(* Logix 5000 project; controller _1407974_PSG_7315 vendor 1 type 14 code 154 rev 20.11; software revision 20.06 *)
// S/O:1407974
// MODEL: PSG P7315

TASK MainTask (continuous, watchdog 500 ms) : MainProgram

MODULES
   Local : vendor 1 type 14 code 154 (PointIO 0, rev 20.11)
      Delta_V : 1756-ENBT (Ethernet 192.168.1.1, rev 3.1)
      Remote : vendor 1 type 12 code 132 (Ethernet 192.168.1.51, rev 4.10, Output RPI 20 ms)
         RTD_In_Module : vendor 1 type 115 code 125 (ArmorPoint 2, rev 3.4, Input RPI 50 ms)
         DI_1_Module : vendor 1 type 7 code 201 (ArmorPoint 1, rev 3.22, Input RPI 50 ms)
         DO_Module : vendor 1 type 7 code 209 (ArmorPoint 3, rev 3.22, Output RPI 50 ms)
         AO_Module : vendor 1 type 115 code 127 (ArmorPoint 4, rev 3.4, Output RPI 80 ms)
      Local_AI_Slot_2 : 1734-IE2C (PointIO 2, rev 3.1, Input RPI 80 ms)
       : vendor 1 type 115 code 211 (PointIO 3, rev 3.1, Output RPI 80 ms)
      Discrete_IO : Embedded (PointIO 1, rev 20.11, Output RPI 20 ms)
END_MODULES

TYPE Analog_Input :
STRUCT
   Raw : REAL;
   Scaled : REAL;
   Fault : BOOL;
   Under_Range : BOOL;
   Over_Range : BOOL;
   Control_Set_Point : REAL;
   Alarm_Low_Set_Point : REAL;
   Alarm_High_Set_Point : REAL;
   Temp_Set_Point : REAL;
   Tieback : REAL;
   SCP : SCP;
   EU_Low : REAL;
   EU_hi : REAL;
   PID : PID;
   Low_Stpt : REAL;
   Low_Low_Stpt : REAL;
   High_Stpt : REAL;
   High_High_Stpt : REAL;
   Ana_Out : Analog_Output;
END_STRUCT
END_TYPE

TYPE Analog_Output :
STRUCT
   Scaled : REAL;
   Manual : REAL;
   Fault : BOOL;
   Raw : REAL;
   SCP : SCP;
   ManSCP : SCP;
   Set_Point_Entry : OIT_Set_Point_Entry;
END_STRUCT
END_TYPE

TYPE AW :
STRUCT
   Network_Ack : INT[2];
   Network_Ack_ONS : INT[2];
   Network_Ack_Handshake : INT[2];
   Network_Ack_Latch : INT[2];
   Network_Ack_All_Latch : BOOL;
   Remote_Ack_All : INT;
   Network_Alarm_Ack : INT[2];
   OIT_Ack : INT[2];
   Latch_Bit : INT[2];
   Ack : INT[2];
   No_Active_Alarms : BOOL;
   No_Active_Warnings : BOOL;
   Silence : INT[2];
   All_Alarms_Acknowledged : BOOL;
   All_Warnings_Acknowledged : BOOL;
   Alarms_Silenced : BOOL;
   Warnings_Silenced : BOOL;
   OIT_Silence_PB : Push_Button;
   Alarm_Silence_Latch : BOOL;
   Warning_Silence_Latch : BOOL;
END_STRUCT
END_TYPE

TYPE Date_Time :
STRUCT
   Set_Push_Button : BOOL;
   Handshake : BOOL;
END_STRUCT
END_TYPE

TYPE Discrete_Out :
STRUCT
   Activate : BOOL;
   Maint_Latch : Latched_Push_Button;
END_STRUCT
END_TYPE

TYPE OIT_Connections :
STRUCT
   Current_Minute : DINT;
   Update : BOOL;
   Current_Screen : DINT;
   Previous_Minute : DINT;
END_STRUCT
END_TYPE

TYPE OIT_Message :
STRUCT
   Operational_Mode : INT;
   Operational_Step_State : INT;
   Information_Message_Number : INT;
   Feed_Water_Pump_Status : INT;
   Low_Level_Swtitch_Status : INT;
   Hi_Hi_Level_Switch_Status : INT;
   Pure_Steam_Temp_Status : INT;
   Pure_Steam_Conductivity_Status : INT;
   Alarm_Warning_Status : INT;
END_STRUCT
END_TYPE

TYPE OIT_Popup :
STRUCT
   Call : BOOL;
   Called : BOOL;
   Timer : TIMER;
   Close : BOOL;
END_STRUCT
END_TYPE

TYPE OIT_Set_Point_Entry :
STRUCT
   OIT_Enter : Push_Button;
   OIT_Set_Point_Buffer : REAL;
END_STRUCT
END_TYPE

TYPE Push_Button :
STRUCT
   Push_Button : BOOL;
   Indicator : BOOL;
   One_Shot : BOOL;
   Handshake : BOOL;
END_STRUCT
END_TYPE

TYPE Unit_Status :
STRUCT
   ON : BOOL;
   OFF : BOOL;
   READY : BOOL;
   FILLING : BOOL;
   HEATING : BOOL;
   RUNNING : BOOL;
   COOLING : BOOL;
   MAINTENANCE : BOOL;
END_STRUCT
END_TYPE

ADD_ON_INSTRUCTION Latched_Push_Button   (* revision 1.0 *)
VAR_INPUT
   OIT_Momentary_PB : BOOL; {required}
END_VAR
VAR_OUTPUT
   OIT_Status : BOOL; {access Read Only, required}
END_VAR
VAR
   OIT_Toggle_ONS : BOOL;
   OIT_Select_ONS : BOOL;
END_VAR

ROUTINE Logic   (* ladder *)
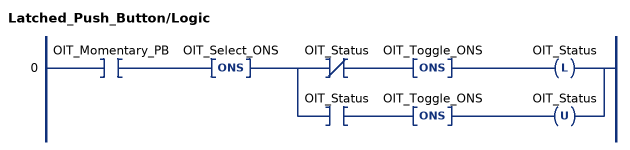
   0: XIC(OIT_Momentary_PB)ONS(OIT_Select_ONS)[XIO(OIT_Status) ONS(OIT_Toggle_ONS) OTL(OIT_Status) ,XIC(OIT_Status) ONS(OIT_Toggle_ONS) OTU(OIT_Status) ];
END_ROUTINE
END_ADD_ON_INSTRUCTION

ADD_ON_INSTRUCTION SCP   (* revision 1.0, vendor Rockwell Automation *)
VAR_INPUT
   Input : REAL; {required}
   InputMin : REAL; {required}
   InputMax : REAL; {required}
   ScaledMin : REAL; {required}
   ScaledMax : REAL; {required}
END_VAR
VAR_OUTPUT
   Output : REAL; {access Read Only, required}
END_VAR
VAR
   Temp4 : REAL;
   Temp3 : REAL;
   Temp2 : REAL;
   Temp1 : REAL;
   Offset : REAL;
   Rate : REAL;
   Out : REAL;
END_VAR

ROUTINE Logic   (* ladder *)
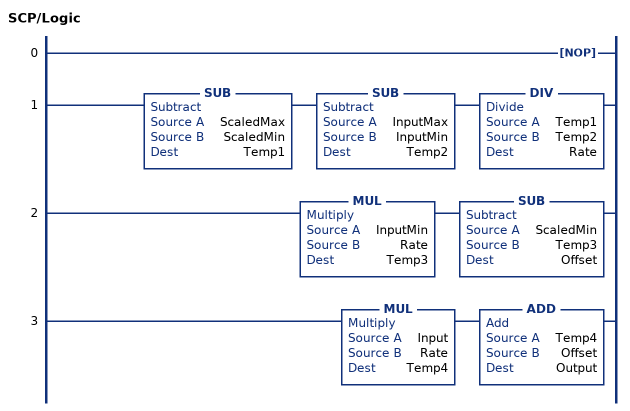
   0: NOP();
   1: SUB(ScaledMax,ScaledMin,Temp1)SUB(InputMax,InputMin,Temp2)DIV(Temp1,Temp2,Rate);
   2: MUL(InputMin,Rate,Temp3)SUB(ScaledMin,Temp3,Offset);
   3: MUL(Input,Rate,Temp4)ADD(Temp4,Offset,Output);
END_ROUTINE
END_ADD_ON_INSTRUCTION

VAR_GLOBAL   (* controller tags *)
   AI_L_2_0_Pure_Steam_Conductivity : Analog_Input := (Raw := 9171.0, Scaled := 0.8994354, Alarm_High_Set_Point := 1.2, SCP.Input := 9171.0, SCP.InputMin := 3277.0, SCP.InputMax := 16383.0, SCP.ScaledMax := 2.0, SCP.Output := 0.8994354);
   AI_L_2_1_FW_Press_Low_Warning : OIT_Set_Point_Entry := (OIT_Set_Point_Buffer := 5.0);
   AI_L_2_1_FW_Pressure : Analog_Input := (Raw := 3321.0, Scaled := 0.5035858, Control_Set_Point := 80.0, Alarm_High_Set_Point := 2.0, Temp_Set_Point := 80.0, SCP.Input := 3321.0, SCP.InputMin := 3277.0, SCP.InputMax := 16383.0, SCP.ScaledMax := 150.0, SCP.Output := 0.5035858, Low_Stpt := 5.0);
   AI_R_2_0_Pure_Steam_Temperature : Analog_Input := (Scaled := 139.6, Control_Set_Point := 140.0, Alarm_Low_Set_Point := 102.0, Alarm_High_Set_Point := 176.0, Temp_Set_Point := 140.0);
   AI_R_2_1_Cond_Pure_Steam_Temperature : Analog_Input := (Scaled := 99.9, Alarm_High_Set_Point := 99.0);
   Alarm_Emergency_Stop : ALIAS FOR Alarms_Warnings.Latch_Bit[0].0;
   Alarm_Emergency_Stop_Ack : ALIAS FOR Alarms_Warnings.Ack[0].0;
   Alarm_Pure_Steam_High_Temp_Timer : TIMER := (PRE := 60000);
   Alarm_Pure_Steam_High_Temperature : ALIAS FOR Alarms_Warnings.Latch_Bit[0].4;
   Alarm_Pure_Steam_High_Temperature_Ack : ALIAS FOR Alarms_Warnings.Ack[0].4;
   Alarm_Pure_Steam_Temp_Error_Timer : TIMER := (PRE := 5000);
   Alarm_Pure_Steam_Temp_Input_Error : ALIAS FOR Alarms_Warnings.Latch_Bit[0].5;
   Alarm_Pure_Steam_Temp_Input_Error_Ack : ALIAS FOR Alarms_Warnings.Ack[0].5;
   Alarm_Rupture_Disk_Failure : ALIAS FOR Alarms_Warnings.Latch_Bit[0].1;
   Alarm_Rupture_Disk_Failure_Timer : TIMER := (PRE := 750);
   Alarm_Rupture_Disk_Faiure_Ack : ALIAS FOR Alarms_Warnings.Ack[0].1;
   Alarm_Separator_High_Level : ALIAS FOR Alarms_Warnings.Latch_Bit[0].2;
   Alarm_Separator_High_Level_Ack : ALIAS FOR Alarms_Warnings.Ack[0].2;
   Alarm_Separator_High_Level_Timer : TIMER := (PRE := 120000);
   Alarm_Separator_Low_Level : ALIAS FOR Alarms_Warnings.Latch_Bit[0].3;
   Alarm_Separator_Low_Level_Ack : ALIAS FOR Alarms_Warnings.Ack[0].3;
   Alarm_Separator_Low_Level_Timer_A : TIMER := (PRE := 600000);
   Alarm_Separator_Low_Level_Timer_B : TIMER := (PRE := 60000);
   Alarms_Warnings : AW := (Network_Ack[1] := 32, Network_Ack_Handshake[0] := 1, Network_Ack_Handshake[1] := 1, Latch_Bit[1] := 2#0000_0000_0000_0001, No_Active_Alarms := 1, All_Alarms_Acknowledged := 1, Alarms_Silenced := 1);
   AO_L_3_0_VFD_SPEED : Analog_Output := (Scaled := 100.0, Manual := 100.0, Raw := 100.0);
   AO_L_3_1_Available : Analog_Output := (SCP.InputMax := 100.0, SCP.ScaledMin := 3277.0, SCP.ScaledMax := 16383.0, SCP.Output := 3277.0, ManSCP.InputMax := 100.0, ManSCP.ScaledMin := 3277.0, ManSCP.ScaledMax := 16383.0, ManSCP.Output := 3277.0);
   AO_L_3_2_Available : Analog_Output := (SCP.InputMax := 100.0, SCP.ScaledMin := 3277.0, SCP.ScaledMax := 16383.0, SCP.Output := 3277.0, ManSCP.InputMax := 100.0, ManSCP.ScaledMin := 3277.0, ManSCP.ScaledMax := 16383.0, ManSCP.Output := 3277.0);
   AO_L_3_3_Available : Analog_Output := (SCP.InputMax := 100.0, SCP.ScaledMin := 3277.0, SCP.ScaledMax := 16383.0, SCP.Output := 3277.0, ManSCP.InputMax := 100.0, ManSCP.ScaledMin := 3277.0, ManSCP.ScaledMax := 16383.0, ManSCP.Output := 3277.0);
   AO_R_4_0_Pure_Steam_Temperature : Analog_Output := (Raw := 54.780636);
   AO_R_4_1_Available : Analog_Output := (SCP.InputMax := 100.0, SCP.ScaledMax := 16383.0, ManSCP.InputMax := 100.0, ManSCP.ScaledMin := 3277.0, ManSCP.ScaledMax := 16383.0, ManSCP.Output := 3277.0);
   Calculated_CV_Max_Value : REAL := 100.0;
   Clean_Steam_Gen_Binary_Data : INT := 8;
   Clean_Steam_Gen_Data : REAL[2] := ([0] := 22.3, [1] := 0.32427895);
   Clean_Steam_Gen_Data3 : INT := 8;
   Cond_Pure_Steam_Conductivity_High : BOOL;
   Cond_Pure_Steam_Hi_Cond_Set_Point_Entry : OIT_Set_Point_Entry := (OIT_Set_Point_Buffer := 1.2);
   Cond_Pure_Steam_Hi_Temp_Set_Point_Entry : OIT_Set_Point_Entry := (OIT_Set_Point_Buffer := 99.0);
   Cond_Pure_Steam_Quality_OK_Latch : BOOL;
   Condensed_Pure_Steam_Warrnings_Disabled : Latched_Push_Button := (OIT_Status := 1);
   Conductivity_Analzyer_Warmup_Delay_Timer : TIMER := (PRE := 600000);
   Cooling_State_Latch_Timer : TIMER := (PRE := 30000, EN := 1, DN := 1);
   Cooling_Status_Debounce_Timer : TIMER := (PRE := 5000);
   DI_L_1_0_Emergency_Stop_Relay : ALIAS FOR DI_Local_1.0;
   DI_L_1_10_Available : ALIAS FOR DI_Local_1.10;
   DI_L_1_11_Available : ALIAS FOR DI_Local_1.11;
   DI_L_1_12_Available : ALIAS FOR DI_Local_1.12;
   DI_L_1_13_Available : ALIAS FOR DI_Local_1.13;
   DI_L_1_14_Feed_Water_Pump_Auto : ALIAS FOR DI_Local_1.14;
   DI_L_1_15_Feed_Water_Pump_Manual : ALIAS FOR DI_Local_1.15;
   DI_L_1_1_Feed_Water_Pump_Aux : ALIAS FOR DI_Local_1.1;
   DI_L_1_2_Pure_Steam_Analyzer_Fault : ALIAS FOR DI_Local_1.2;
   DI_L_1_3_Feed_Water_Analyzer_Fault : ALIAS FOR DI_Local_1.3;
   DI_L_1_4_Available : ALIAS FOR DI_Local_1.4;
   DI_L_1_5_Available : ALIAS FOR DI_Local_1.5;
   DI_L_1_6_Available : ALIAS FOR DI_Local_1.6;
   DI_L_1_7_Available : ALIAS FOR DI_Local_1.7;
   DI_L_1_8_Available : ALIAS FOR DI_Local_1.8;
   DI_L_1_9_Available : ALIAS FOR DI_Local_1.9;
   DI_Local_1 : INT := 7;
   DI_R_1_0_Hi_Hi_Level_LSHH_1950 : ALIAS FOR DI_Remote_1.0;
   DI_R_1_1_Hi_Level_LSH_1950 : ALIAS FOR DI_Remote_1.1;
   DI_R_1_2_Mid_Level_LSM_1950 : ALIAS FOR DI_Remote_1.2;
   DI_R_1_3_Low_Level_LSL_1950 : ALIAS FOR DI_Remote_1.3;
   DI_R_1_4_Air_Low_Pressure_PSL_4030 : ALIAS FOR DI_Remote_1.4;
   DI_R_1_5_Burst_Disk_Sensor_PSH_5820 : ALIAS FOR DI_Remote_1.5;
   DI_R_1_6_Available : ALIAS FOR DI_Remote_1.6;
   DI_R_1_7_Available : ALIAS FOR DI_Remote_1.7;
   DI_Remote_1 : INT := 59;
   DO_L_1_0_Alarm_Relay_Coil : Discrete_Out;
   DO_L_1_0_Alarm_Relay_Out : BOOL;
   DO_L_1_10_Available : Discrete_Out;
   DO_L_1_10_Spare_Out : BOOL;
   DO_L_1_11_Available : Discrete_Out;
   DO_L_1_11_Spare_Out : BOOL;
   DO_L_1_12_Available : Discrete_Out;
   DO_L_1_12_Spare_Out : BOOL;
   DO_L_1_13_Available : Discrete_Out;
   DO_L_1_13_Spare_Out : BOOL;
   DO_L_1_13_VFD_Relay_In : BOOL;
   DO_L_1_14_Feed_Pump_Out : BOOL;
   DO_L_1_14_Feed_Water_Pump_Contactor : Discrete_Out;
   DO_L_1_15_Feed_Pump_Light_Out : BOOL;
   DO_L_1_15_Feed_Water_Pump_On_Light : Discrete_Out;
   DO_L_1_1_Alarm_Horn : Discrete_Out := (Activate := 1);
   DO_L_1_1_Alarm_Horn_Out : BOOL := 1;
   DO_L_1_2_Alarm_Light : Discrete_Out := (Activate := 1);
   DO_L_1_2_Alarm_Light_Out : BOOL := 1;
   DO_L_1_3_Ready_Light : Discrete_Out;
   DO_L_1_3_Ready_Light_Out : BOOL;
   DO_L_1_4_Running_Light : Discrete_Out;
   DO_L_1_4_Running_Light_Out : BOOL;
   DO_L_1_5_Hour_Meter : Discrete_Out;
   DO_L_1_5_Hour_Meter_Out : BOOL;
   DO_L_1_6_Available : Discrete_Out;
   DO_L_1_6_Spare_Out : BOOL;
   DO_L_1_7_Available : Discrete_Out;
   DO_L_1_7_Spare_Out : BOOL;
   DO_L_1_8_Available : Discrete_Out;
   DO_L_1_8_Spare_Out : BOOL;
   DO_L_1_9_Available : Discrete_Out;
   DO_L_1_9_Spare_Out : BOOL;
   DO_Local_1 : INT := 6;
   DO_R_3_0_Pure_Steam_Control_Valve_Out : BOOL;
   DO_R_3_0_Pure_Steam_Temp_Control_YV_4110 : Discrete_Out;
   DO_R_3_1_Pri_Level_Valve_Out : BOOL;
   DO_R_3_1_Primary_Level_Control_YV_4760 : Discrete_Out;
   DO_R_3_2_Sec_Level_Valve_Out : BOOL;
   DO_R_3_2_Secondary_Level_Control_YV_4770 : Discrete_Out;
   DO_R_3_3_Coolant_Shutoff_FCV_3025 : Discrete_Out;
   DO_R_3_3_Coolant_Valve_Out : BOOL;
   DO_R_3_4_Degasser_Vent_Out : BOOL := 1;
   DO_R_3_4_Degasser_Vent_YV_4255 : Discrete_Out := (Activate := 1);
   DO_R_3_5_FDW_TR : Discrete_Out;
   DO_R_3_5_Spare_Out : BOOL;
   DO_R_3_6_Available : Discrete_Out;
   DO_R_3_6_Spare_Out : BOOL;
   DO_R_3_7_Available : Discrete_Out;
   DO_R_3_7_Spare_Out : BOOL;
   DO_Remote_3 : INT := 16;
   F8_0_9 : REAL[10] := ([0] := 139.6, [1] := 0.8994354); {produced, access Read Only}
   F8_50_59 : REAL[10]; {produced}
   Feed_Water_Conductivity_High : BOOL;
   Feed_Water_Pressure_Set_Point_Entry : OIT_Set_Point_Entry := (OIT_Set_Point_Buffer := 80.0);
   Feed_Water_Pump_Delay_Timer : TIMER := (PRE := 3000);
   Feedwater_Pressure_PID : PID := (CTL := 37504, INI := 1, OLH := 1, DVPA := 1, PVHA := 1, SP := 80.0, KP := 5.5, KI := 0.5, KD := 0.06, MAXS := 4095.0, SO := 100.0, MAXO := 100.0, UPD := 0.44, PV := 0.5035858, ERR := 79.496414, OUT := 100.0, MAXI := 4095.0, TIE := 2.4420025, MAXTIE := 4095.0, DATA[0] := 96.912155, DATA[1] := -0.19676125, DATA[2] := 0.5035858, DATA[3] := 79.496414, DATA[4] := 80.0, DATA[5] := 0.024420025, DATA[6] := 1.0, DATA[7] := 7.1, DATA[8] := 5.5, DATA[9] := 0.5, DATA[10] := 0.06, DATA[11] := 5.5, DATA[12] := 0.5, DATA[13] := 0.06, DATA[16] := 0.024420025);
   Feedwater_Pressure_PID_Auto_Mode : Push_Button := (One_Shot := 1);
   Feedwater_Pressure_PID_Manual_Mode : Push_Button;
   Free_Run_Pulse_Timer : TIMER := (PRE := 2048, ACC := 1145, EN := 1, TT := 1);
   FW_Cond_Analyzer_Return_Delay : TIMER := (PRE := 10000, ACC := 10000, EN := 1, DN := 1);
   FW_Press_PID_Gain_Set_Point_Entry : OIT_Set_Point_Entry := (OIT_Set_Point_Buffer := 5.5);
   FW_Press_PID_Manual_Output_Entry : OIT_Set_Point_Entry := (OIT_Set_Point_Buffer := 50.0);
   FW_Press_PID_Rate_Set_Point_Entry : OIT_Set_Point_Entry := (OIT_Set_Point_Buffer := 0.06);
   FW_Press_PID_Reset_SetPoint_Entry : OIT_Set_Point_Entry := (OIT_Set_Point_Buffer := 0.5);
   FW_Press_PID_Temp_Set_Point_Entry : OIT_Set_Point_Entry := (OIT_Set_Point_Buffer := 150.0);
   Lamp_Test : Push_Button;
   Local_Remote : Latched_Push_Button;
   Login_Popup : OIT_Popup := (Timer.PRE := 30000);
   Login_Required_Popup : OIT_Popup := (Timer.PRE := 30000);
   Low_Feedwater_Pressure : BOOL;
   Low_Level_Latch : BOOL;
   Maintenance_Mode : Latched_Push_Button;
   Maintenance_Screen_Not_Displayed : BOOL;
   N7_0_9 : INT[10] := ([0] := 40, [1] := 8210); {produced, access Read Only}
   N7_100_109 : INT[10] := ([0] := 26, [1] := 1); {produced}
   Network_Ack_All : BOOL;
   Network_AI_L_2_0_Pure_Steam_Conductivity : REAL := 0.8994354;
   Network_AI_L_2_1_Feedwater_Pressure : REAL := 0.5035858;
   Network_AI_L_2_1_FW_Pressure_Scaled : DINT := 1;
   Network_AI_R_2_0_Pure_Steam_Temperature : REAL := 139.6;
   Network_AI_R_2_1_Cond_Pure_Steam_Temp : REAL := 99.9;
   Network_AO_R_4_0_Pure_Steam_Man_Control : REAL;
   Network_AO_R_4_0_Pure_Steam_Temp_Control : REAL;
   Network_AO_R_4_1_Available_Manual : REAL;
   Network_AO_R_4_1_Available_Scaled : REAL;
   Network_Cond_PS_Temp_High_Set_Point : REAL := 99.0;
   Network_DI_Local_1 : INT := 7;
   Network_DI_Remote_1 : INT := 59;
   Network_DO_Local_1 : INT := 6;
   Network_DO_Remote_3 : INT := 16;
   Network_Feedwater_Pressure_PID : DINT;
   Network_Feedwater_Pressure_PID_KD : DINT;
   Network_Feedwater_Pressure_PID_KI : DINT;
   Network_Feedwater_Pressure_PID_KP : DINT := 6;
   Network_Feedwater_Pressure_PID_SP : DINT := 80;
   Network_FW_Low_Pressure_Warning_SP : DINT := 5;
   Network_Input_Ack_All : BOOL;
   Network_Input_Silence : BOOL;
   Network_Input_Silence_ONS : BOOL;
   Network_Input_Start : BOOL;
   Network_Input_Start_ONS : BOOL;
   Network_Input_Stop : BOOL;
   Network_Input_Stop_ONS : BOOL;
   Network_PID_Ramp_Time_Seconds : DINT := 120;
   Network_Pure_Steam_Conductivity_SetPoint : REAL := 1.2;
   Network_Pure_Steam_Temp_High_Set_Point : REAL := 176.0;
   Network_Pure_Steam_Temp_Lo_Set_Point : REAL := 102.0;
   Network_Pure_Steam_Temp_PID_Gain : REAL := 3.75;
   Network_Pure_Steam_Temp_PID_Rate : REAL := 0.05;
   Network_Pure_Steam_Temp_PID_Reset : REAL := 0.05;
   Network_Pure_Steam_Temperature_Set_Point : REAL := 140.0;
   Network_Pure_Steam_Temporary_Set_Point : REAL := 140.0;
   Network_Silence : BOOL;
   Network_Start : BOOL;
   Network_Status_Local_Remote : BOOL;
   Network_Status_Maintenance_Mode : BOOL;
   Network_Status_No_Active_Alarms : BOOL := 1;
   Network_Status_No_Active_Warnings : BOOL;
   Network_Status_Unit_Cooling : BOOL := 1;
   Network_Status_Unit_Filling : BOOL;
   Network_Status_Unit_Heating : BOOL;
   Network_Status_Unit_OFF : BOOL := 1;
   Network_Status_Unit_ON : BOOL;
   Network_Status_Unit_Ready : BOOL;
   Network_Status_Unit_Running : BOOL;
   Network_Stop : BOOL;
   Netwrok_Input_Ack_All_ONS : BOOL;
   OIT : OIT_Connections := (Current_Minute := 19, Current_Screen := 2, Previous_Minute := 19);
   OIT_Auto_Time_Date_Sync : TIMER := (PRE := 2000);
   OIT_Auto_Time_Date_Sync_Interval : TIMER := (PRE := 600000, ACC := 485432, EN := 1, TT := 1);
   OIT_Day_Set : Push_Button;
   OIT_Hour_Set : Push_Button;
   OIT_Message : OIT_Message := (Operational_Step_State := 4, Low_Level_Swtitch_Status := 1, Hi_Hi_Level_Switch_Status := 1, Alarm_Warning_Status := 1);
   OIT_Message_FW_Cond_Status : DINT;
   OIT_Minute_Set : Push_Button;
   OIT_Month_Set : Push_Button;
   OIT_SPEED_COMMAND : REAL := 85.0;
   OIT_Year_Set : Push_Button;
   PID_Auto_Mode : Push_Button := (One_Shot := 1);
   PID_CV_Max_Value_Initialize : BOOL;
   PID_Loop_Trigger_Timer : TIMER := (PRE := 100, ACC := 31, EN := 1, TT := 1);
   PID_Manual_Mode : Push_Button;
   PID_Ramp_Time_Seconds : DINT := 120;
   PID_Ramp_Timer : TIMER := (PRE := 120000);
   Primary_Feed_Water_Valve_Open_Timer : TIMER := (PRE := 55000, ACC := 7557, EN := 1, TT := 1);
   PS_Temp_GEQ_SetPoint_Minus_5_Deg : BOOL;
   PS_Temp_Setpoint_Minus_5_Deg : REAL := 135.0;
   Pulse_Bit : BOOL := 1;
   Pure_Steam_High_Temp_Set_Point_Entry : OIT_Set_Point_Entry := (OIT_Set_Point_Buffer := 176.0);
   Pure_Steam_Low_Temp_Set_Point_Entry : OIT_Set_Point_Entry := (OIT_Set_Point_Buffer := 102.0);
   Pure_Steam_Temp_Cntrl_Output_SCP : SCP := (InputMax := 100.0, ScaledMin := 3277.0, ScaledMax := 16383.0, Output := 3277.0);
   Pure_Steam_Temp_Manual_Output_SCP : SCP := (InputMax := 100.0, ScaledMin := 3277.0, ScaledMax := 16383.0, Output := 3277.0);
   Pure_Steam_Temp_Output_Clamp : BOOL := 1;
   Pure_Steam_Temp_PID_Gain_Set_Point_Entry : OIT_Set_Point_Entry := (OIT_Set_Point_Buffer := 3.75);
   Pure_Steam_Temp_PID_Manual_Output_Entry : OIT_Set_Point_Entry;
   Pure_Steam_Temp_PID_Ramp_Time_Entry : OIT_Set_Point_Entry := (OIT_Set_Point_Buffer := 120.0);
   Pure_Steam_Temp_PID_Rate_Set_Point_Entry : OIT_Set_Point_Entry := (OIT_Set_Point_Buffer := 0.05);
   Pure_Steam_Temp_PID_Reset_SetPoint_Entry : OIT_Set_Point_Entry := (OIT_Set_Point_Buffer := 0.05);
   Pure_Steam_Temp_PID_Temp_Set_Point_Entry : OIT_Set_Point_Entry := (OIT_Set_Point_Buffer := 138.0);
   Pure_Steam_Temperature : PID := (CTL := 33408, INI := 1, DVPA := 1, PVHA := 1, SP := 140.0, KP := 3.75, KI := 0.05, KD := 0.05, MAXS := 176.0, SO := 54.780636, MAXO := 100.0, UPD := 0.05, PV := 139.6, ERR := 0.3999939, OUT := 54.780636, MAXI := 176.0, TIE := 54.780067, MAXCV := 100.0, MAXTIE := 100.0, DATA[0] := 53.928375, DATA[1] := -1269.091, DATA[2] := 139.6, DATA[3] := 0.3999939, DATA[4] := 140.0, DATA[5] := 0.5681818, DATA[6] := 1.0, DATA[7] := 0.85, DATA[8] := 3.75, DATA[9] := 0.05, DATA[10] := 0.05, DATA[11] := 3.75, DATA[12] := 0.05, DATA[13] := 0.05, DATA[15] := 1.0, DATA[16] := 1.0);
   Pure_Steam_Temperature_Set_Point_Entry : OIT_Set_Point_Entry := (OIT_Set_Point_Buffer := 140.0);
   Read_PLC_Clock : DINT[7] := ([0] := 2026, [1] := 9, [2] := 22, [3] := 9, [4] := 46, [5] := 41, [6] := 18779);
   Set_PLC_Clock : DINT[7] := ([0] := 2019, [1] := 8, [2] := 26, [3] := 7, [4] := 47);
   Start : Push_Button;
   Start_Stop_Popup : OIT_Popup := (Timer.PRE := 30000);
   Stop : Push_Button;
   Unit_Hot : BOOL := 1;
   Unit_Status : Unit_Status := (OFF := 1, COOLING := 1);
   VFD_HANDS_REFERENCE_SPEED : SCP := (Input := 85.0, InputMax := 100.0, ScaledMin := 1638.0, ScaledMax := 8191.0, Output := 7208.05);
   VFD_Relay_Input : BOOL;
   VFD_Speed_Cntrl_Output_SCP : Analog_Output;
   VFD_Speed_Control_Auto : SCP := (Input := 100.0, InputMax := 100.0, ScaledMin := 1638.0, ScaledMax := 8191.0, Output := 8191.0);
   VFD_SPEED_CONTROL_MANUAL : SCP := (Input := 100.0, InputMax := 100.0, ScaledMin := 1638.0, ScaledMax := 8191.0, Output := 8191.0);
   Warning_Air_Low_Pressure_Timer : TIMER := (PRE := 60000);
   Warning_Cond_Pure_Steam_Analyzer_Fault : ALIAS FOR Alarms_Warnings.Latch_Bit[1].4;
   Warning_Cond_Pure_Steam_Analyzer_Timer : TIMER := (PRE := 5000);
   Warning_Cond_Pure_Steam_Anlzr_Fault_Ack : ALIAS FOR Alarms_Warnings.Ack[1].4;
   Warning_Cond_Pure_Steam_Conduct_Timer : TIMER := (PRE := 10000);
   Warning_Cond_Pure_Steam_Conductivity : ALIAS FOR Alarms_Warnings.Latch_Bit[1].3;
   Warning_Cond_Pure_Steam_Conductivity_Ack : ALIAS FOR Alarms_Warnings.Ack[1].3;
   Warning_Cond_Pure_Steam_Hi_Temp_Timer : TIMER := (PRE := 30000);
   Warning_Cond_Pure_Steam_High_Temp : ALIAS FOR Alarms_Warnings.Latch_Bit[1].8;
   Warning_Cond_Pure_Steam_High_Temp_Ack : ALIAS FOR Alarms_Warnings.Ack[1].8;
   Warning_Evaporator_Low_Pressure_Ack : ALIAS FOR Alarms_Warnings.Ack[1].5;
   Warning_Evaporator_Low_Pressure_Timer : TIMER := (PRE := 60000);
   Warning_Feed_Water_Analyer_Fault_Ack : ALIAS FOR Alarms_Warnings.Ack[1].6;
   Warning_Feed_Water_Analyzer_Fault : ALIAS FOR Alarms_Warnings.Latch_Bit[1].6;
   Warning_Feed_Water_Analyzer_Timer : TIMER := (PRE := 5000);
   Warning_Feed_Water_Conductivity : ALIAS FOR Alarms_Warnings.Latch_Bit[1].5;
   Warning_Feed_Water_Conductivity_Ack : ALIAS FOR Alarms_Warnings.Ack[1].5;
   Warning_Feed_Water_Conductivity_Timer : TIMER := (PRE := 5000);
   Warning_Feed_Water_Pump_Fault : ALIAS FOR Alarms_Warnings.Latch_Bit[1].1;
   Warning_Feed_Water_Pump_Fault_Ack : ALIAS FOR Alarms_Warnings.Ack[1].1;
   Warning_Feed_Water_Pump_Fault_Timer : TIMER := (PRE := 5000);
   Warning_Feedwater_Low_Pressure : ALIAS FOR Alarms_Warnings.Latch_Bit[1].9;
   Warning_Feedwater_Press_Low_Pressure_Ack : ALIAS FOR Alarms_Warnings.Ack[1].9;
   Warning_FW_Press_Low_Pressure_Timer : TIMER := (PRE := 120000);
   Warning_Instrument_Air_Low_Pressure : ALIAS FOR Alarms_Warnings.Latch_Bit[1].2;
   Warning_Instrument_Air_Low_Pressure_Ack : ALIAS FOR Alarms_Warnings.Ack[1].2;
   Warning_Plant_Steam_Low_Pressure_Ack : ALIAS FOR Alarms_Warnings.Ack[1].4;
   Warning_Plant_Steam_Low_Pressure_Timer : TIMER := (PRE := 60000);
   Warning_PLC_OIT_Comm_Counter : COUNTER := (PRE := 2);
   Warning_PLC_OIT_Comm_Timer : TIMER := (PRE := 65000, ACC := 19303, EN := 1, TT := 1);
   Warning_PLC_OIT_Commuications_Ack : ALIAS FOR Alarms_Warnings.Ack[1].0;
   Warning_PLC_OIT_Communications : ALIAS FOR Alarms_Warnings.Latch_Bit[1].0;
   Warning_Pure_Steam_Low_Temp_Timer_A : TIMER := (PRE := 300000);
   Warning_Pure_Steam_Low_Temp_Timer_B : TIMER := (PRE := 120000);
   Warning_Pure_Steam_Low_Temperature : ALIAS FOR Alarms_Warnings.Latch_Bit[1].7;
   Warning_Pure_Steam_Low_Temperature_Ack : ALIAS FOR Alarms_Warnings.Ack[1].7;
END_VAR

PROGRAM MainProgram   (* main routine _010_JSRs *)
VAR
   trial1 : TIMER := (PRE := 1200000, ACC := 208586, EN := 1, TT := 1);
END_VAR

ROUTINE _010_JSRs   (* ladder *)
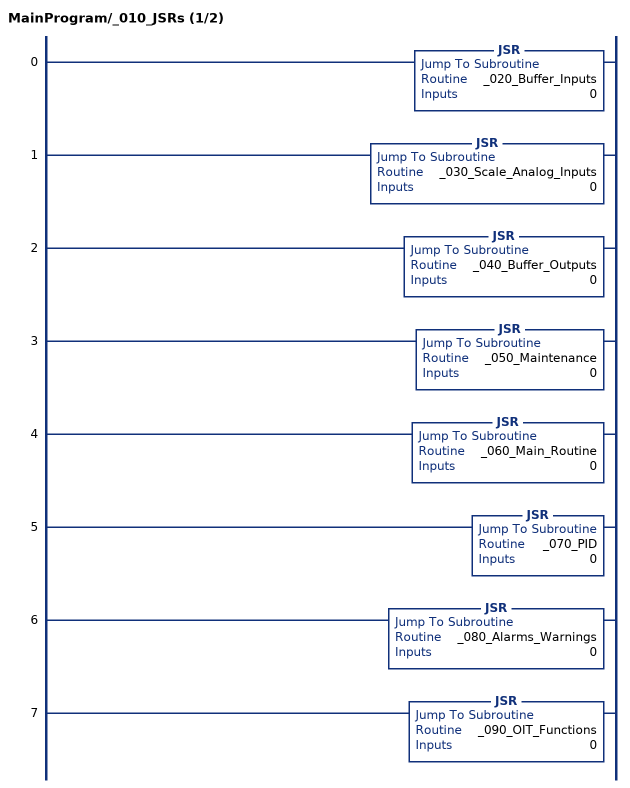
   0: JSR(_020_Buffer_Inputs,0);
   1: JSR(_030_Scale_Analog_Inputs,0);
   2: JSR(_040_Buffer_Outputs,0);
   3: JSR(_050_Maintenance,0);
   4: JSR(_060_Main_Routine,0);
   5: JSR(_070_PID,0);
   6: JSR(_080_Alarms_Warnings,0);
   7: JSR(_090_OIT_Functions,0);
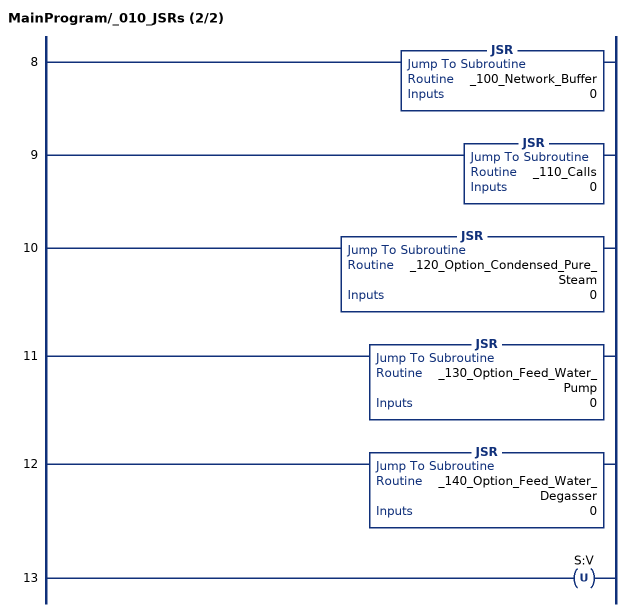
   8: JSR(_100_Network_Buffer,0);
   9: JSR(_110_Calls,0);
   10: JSR(_120_Option_Condensed_Pure_Steam,0);
   11: JSR(_130_Option_Feed_Water_Pump,0);
   12: JSR(_140_Option_Feed_Water_Degasser,0);
   13: OTU(S:V);
END_ROUTINE

ROUTINE _020_Buffer_Inputs   (* ladder *)
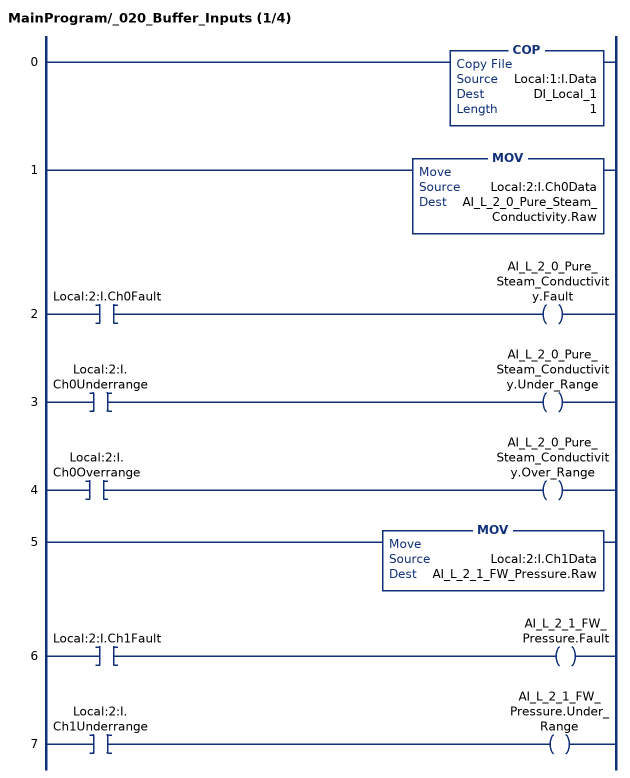
   0: COP(Local:1:I.Data,DI_Local_1,1);
   1: MOV(Local:2:I.Ch0Data,AI_L_2_0_Pure_Steam_Conductivity.Raw);
   2: XIC(Local:2:I.Ch0Fault)OTE(AI_L_2_0_Pure_Steam_Conductivity.Fault);
   3: XIC(Local:2:I.Ch0Underrange)OTE(AI_L_2_0_Pure_Steam_Conductivity.Under_Range);
   4: XIC(Local:2:I.Ch0Overrange)OTE(AI_L_2_0_Pure_Steam_Conductivity.Over_Range);
   5: MOV(Local:2:I.Ch1Data,AI_L_2_1_FW_Pressure.Raw);
   6: XIC(Local:2:I.Ch1Fault)OTE(AI_L_2_1_FW_Pressure.Fault);
   7: XIC(Local:2:I.Ch1Underrange)OTE(AI_L_2_1_FW_Pressure.Under_Range);
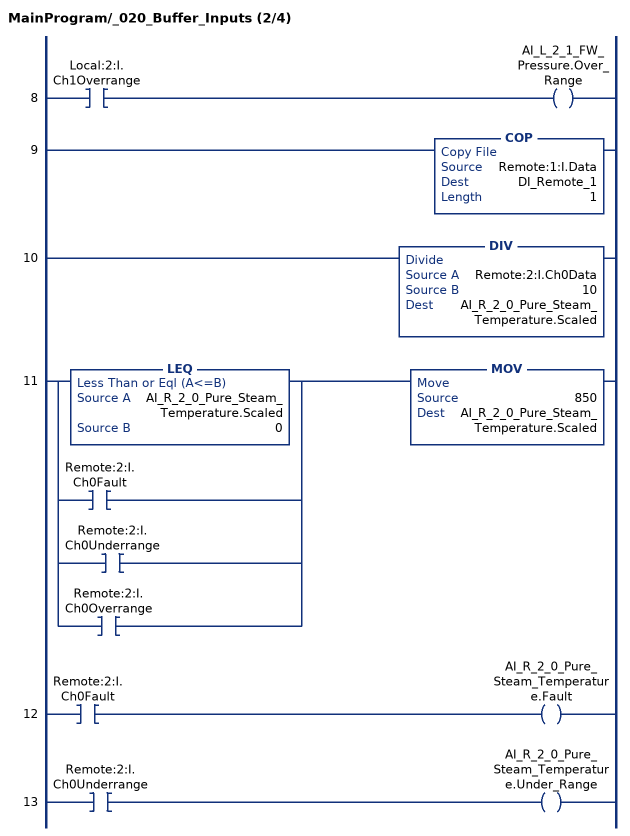
   8: XIC(Local:2:I.Ch1Overrange)OTE(AI_L_2_1_FW_Pressure.Over_Range);
   9: COP(Remote:1:I.Data,DI_Remote_1,1);
   10: DIV(Remote:2:I.Ch0Data,10,AI_R_2_0_Pure_Steam_Temperature.Scaled);
   11: [LEQ(AI_R_2_0_Pure_Steam_Temperature.Scaled,0) ,XIC(Remote:2:I.Ch0Fault) ,XIC(Remote:2:I.Ch0Underrange) ,XIC(Remote:2:I.Ch0Overrange) ]MOV(850,AI_R_2_0_Pure_Steam_Temperature.Scaled);
   12: XIC(Remote:2:I.Ch0Fault)OTE(AI_R_2_0_Pure_Steam_Temperature.Fault);
   13: XIC(Remote:2:I.Ch0Underrange)OTE(AI_R_2_0_Pure_Steam_Temperature.Under_Range);
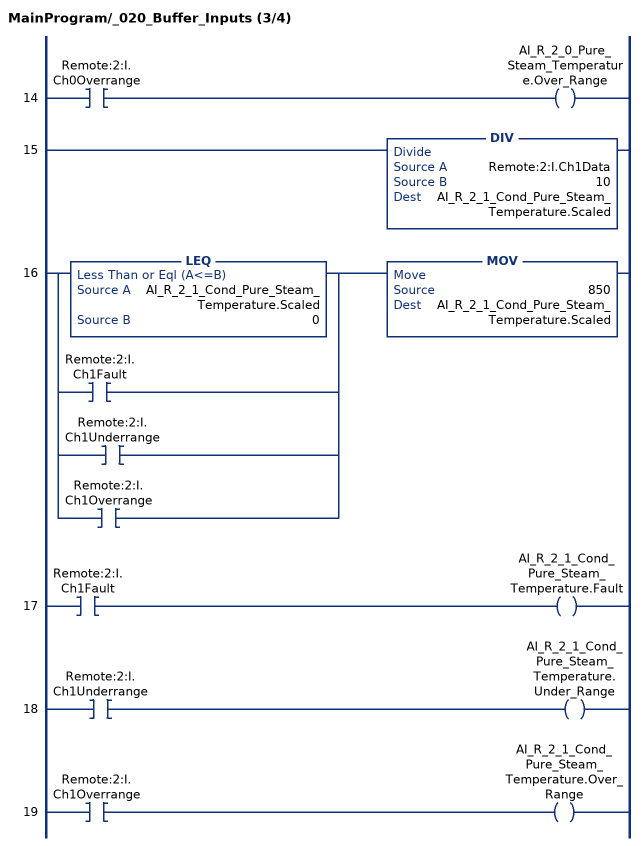
   14: XIC(Remote:2:I.Ch0Overrange)OTE(AI_R_2_0_Pure_Steam_Temperature.Over_Range);
   15: DIV(Remote:2:I.Ch1Data,10,AI_R_2_1_Cond_Pure_Steam_Temperature.Scaled);
   16: [LEQ(AI_R_2_1_Cond_Pure_Steam_Temperature.Scaled,0) ,XIC(Remote:2:I.Ch1Fault) ,XIC(Remote:2:I.Ch1Underrange) ,XIC(Remote:2:I.Ch1Overrange) ]MOV(850,AI_R_2_1_Cond_Pure_Steam_Temperature.Scaled);
   17: XIC(Remote:2:I.Ch1Fault)OTE(AI_R_2_1_Cond_Pure_Steam_Temperature.Fault);
   18: XIC(Remote:2:I.Ch1Underrange)OTE(AI_R_2_1_Cond_Pure_Steam_Temperature.Under_Range);
   19: XIC(Remote:2:I.Ch1Overrange)OTE(AI_R_2_1_Cond_Pure_Steam_Temperature.Over_Range);
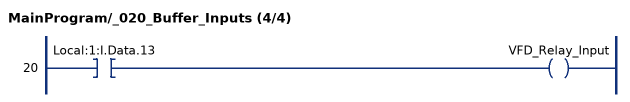
   20: XIC(Local:1:I.Data.13)OTE(VFD_Relay_Input);
END_ROUTINE

ROUTINE _030_Scale_Analog_Inputs   (* ladder *)
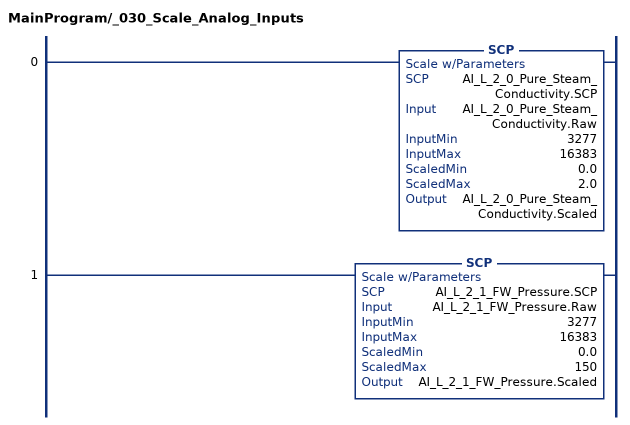
   0: SCP(AI_L_2_0_Pure_Steam_Conductivity.SCP,AI_L_2_0_Pure_Steam_Conductivity.Raw,3277,16383,0.0,2.0,AI_L_2_0_Pure_Steam_Conductivity.Scaled);
   1: SCP(AI_L_2_1_FW_Pressure.SCP,AI_L_2_1_FW_Pressure.Raw,3277,16383,0.0,150,AI_L_2_1_FW_Pressure.Scaled);
END_ROUTINE

ROUTINE _040_Buffer_Outputs   (* ladder *)
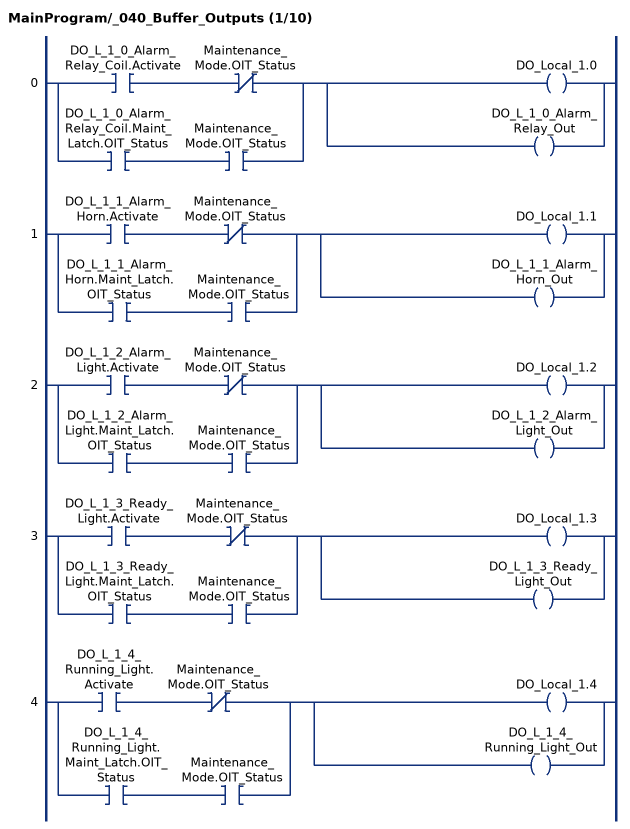
   0: [XIC(DO_L_1_0_Alarm_Relay_Coil.Activate) XIO(Maintenance_Mode.OIT_Status) ,XIC(DO_L_1_0_Alarm_Relay_Coil.Maint_Latch.OIT_Status) XIC(Maintenance_Mode.OIT_Status) ][OTE(DO_Local_1.0) ,OTE(DO_L_1_0_Alarm_Relay_Out) ];
   1: [XIC(DO_L_1_1_Alarm_Horn.Activate) XIO(Maintenance_Mode.OIT_Status) ,XIC(DO_L_1_1_Alarm_Horn.Maint_Latch.OIT_Status) XIC(Maintenance_Mode.OIT_Status) ][OTE(DO_Local_1.1) ,OTE(DO_L_1_1_Alarm_Horn_Out) ];
   2: [XIC(DO_L_1_2_Alarm_Light.Activate) XIO(Maintenance_Mode.OIT_Status) ,XIC(DO_L_1_2_Alarm_Light.Maint_Latch.OIT_Status) XIC(Maintenance_Mode.OIT_Status) ][OTE(DO_Local_1.2) ,OTE(DO_L_1_2_Alarm_Light_Out) ];
   3: [XIC(DO_L_1_3_Ready_Light.Activate) XIO(Maintenance_Mode.OIT_Status) ,XIC(DO_L_1_3_Ready_Light.Maint_Latch.OIT_Status) XIC(Maintenance_Mode.OIT_Status) ][OTE(DO_Local_1.3) ,OTE(DO_L_1_3_Ready_Light_Out) ];
   4: [XIC(DO_L_1_4_Running_Light.Activate) XIO(Maintenance_Mode.OIT_Status) ,XIC(DO_L_1_4_Running_Light.Maint_Latch.OIT_Status) XIC(Maintenance_Mode.OIT_Status) ][OTE(DO_Local_1.4) ,OTE(DO_L_1_4_Running_Light_Out) ];
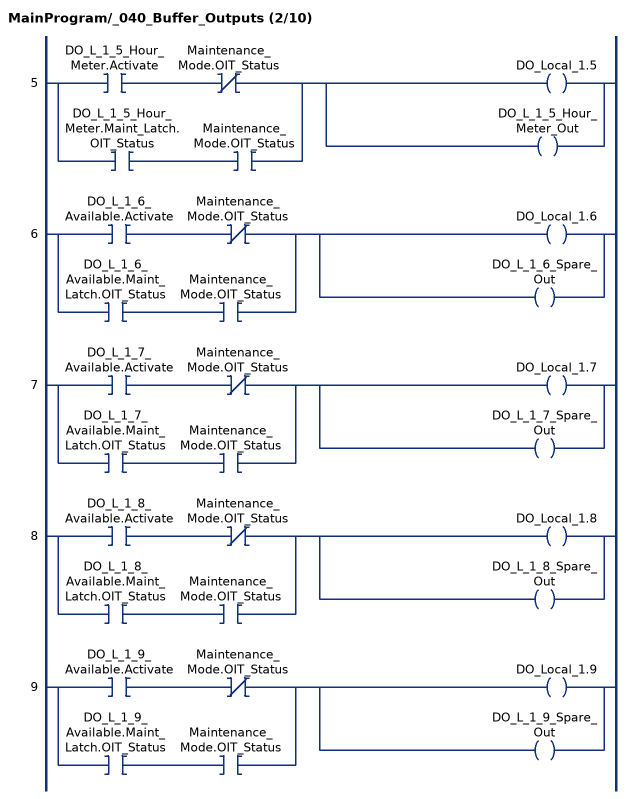
   5: [XIC(DO_L_1_5_Hour_Meter.Activate) XIO(Maintenance_Mode.OIT_Status) ,XIC(DO_L_1_5_Hour_Meter.Maint_Latch.OIT_Status) XIC(Maintenance_Mode.OIT_Status) ][OTE(DO_Local_1.5) ,OTE(DO_L_1_5_Hour_Meter_Out) ];
   6: [XIC(DO_L_1_6_Available.Activate) XIO(Maintenance_Mode.OIT_Status) ,XIC(DO_L_1_6_Available.Maint_Latch.OIT_Status) XIC(Maintenance_Mode.OIT_Status) ][OTE(DO_Local_1.6) ,OTE(DO_L_1_6_Spare_Out) ];
   7: [XIC(DO_L_1_7_Available.Activate) XIO(Maintenance_Mode.OIT_Status) ,XIC(DO_L_1_7_Available.Maint_Latch.OIT_Status) XIC(Maintenance_Mode.OIT_Status) ][OTE(DO_Local_1.7) ,OTE(DO_L_1_7_Spare_Out) ];
   8: [XIC(DO_L_1_8_Available.Activate) XIO(Maintenance_Mode.OIT_Status) ,XIC(DO_L_1_8_Available.Maint_Latch.OIT_Status) XIC(Maintenance_Mode.OIT_Status) ][OTE(DO_Local_1.8) ,OTE(DO_L_1_8_Spare_Out) ];
   9: [XIC(DO_L_1_9_Available.Activate) XIO(Maintenance_Mode.OIT_Status) ,XIC(DO_L_1_9_Available.Maint_Latch.OIT_Status) XIC(Maintenance_Mode.OIT_Status) ][OTE(DO_Local_1.9) ,OTE(DO_L_1_9_Spare_Out) ];
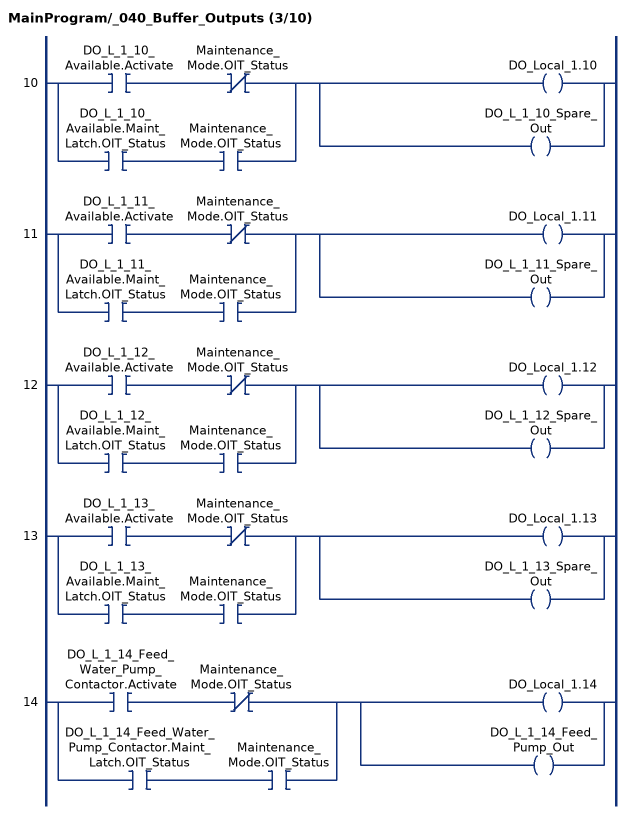
   10: [XIC(DO_L_1_10_Available.Activate) XIO(Maintenance_Mode.OIT_Status) ,XIC(DO_L_1_10_Available.Maint_Latch.OIT_Status) XIC(Maintenance_Mode.OIT_Status) ][OTE(DO_Local_1.10) ,OTE(DO_L_1_10_Spare_Out) ];
   11: [XIC(DO_L_1_11_Available.Activate) XIO(Maintenance_Mode.OIT_Status) ,XIC(DO_L_1_11_Available.Maint_Latch.OIT_Status) XIC(Maintenance_Mode.OIT_Status) ][OTE(DO_Local_1.11) ,OTE(DO_L_1_11_Spare_Out) ];
   12: [XIC(DO_L_1_12_Available.Activate) XIO(Maintenance_Mode.OIT_Status) ,XIC(DO_L_1_12_Available.Maint_Latch.OIT_Status) XIC(Maintenance_Mode.OIT_Status) ][OTE(DO_Local_1.12) ,OTE(DO_L_1_12_Spare_Out) ];
   13: [XIC(DO_L_1_13_Available.Activate) XIO(Maintenance_Mode.OIT_Status) ,XIC(DO_L_1_13_Available.Maint_Latch.OIT_Status) XIC(Maintenance_Mode.OIT_Status) ][OTE(DO_Local_1.13) ,OTE(DO_L_1_13_Spare_Out) ];
   14: [XIC(DO_L_1_14_Feed_Water_Pump_Contactor.Activate) XIO(Maintenance_Mode.OIT_Status) ,XIC(DO_L_1_14_Feed_Water_Pump_Contactor.Maint_Latch.OIT_Status) XIC(Maintenance_Mode.OIT_Status) ][OTE(DO_Local_1.14) ,OTE(DO_L_1_14_Feed_Pump_Out) ];
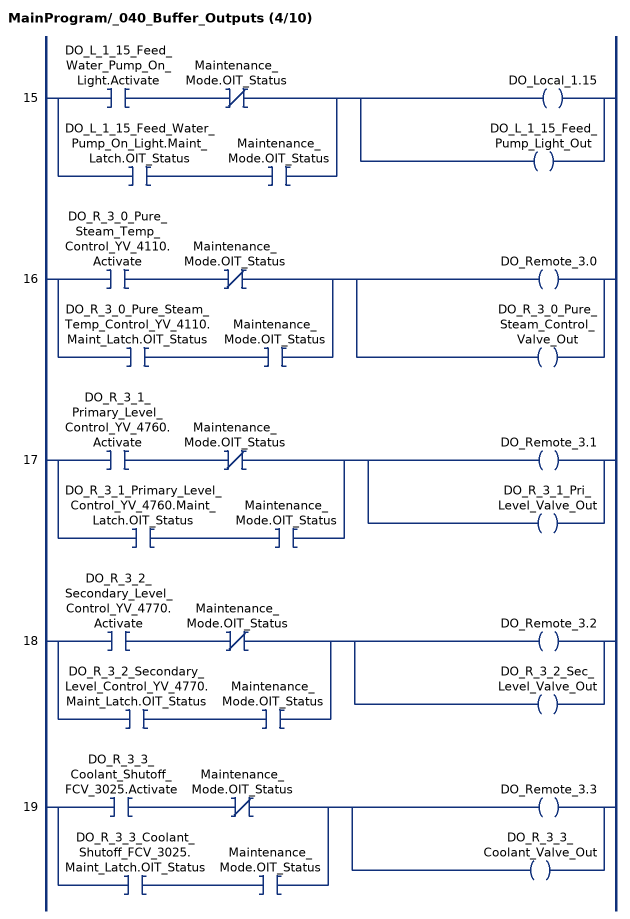
   15: [XIC(DO_L_1_15_Feed_Water_Pump_On_Light.Activate) XIO(Maintenance_Mode.OIT_Status) ,XIC(DO_L_1_15_Feed_Water_Pump_On_Light.Maint_Latch.OIT_Status) XIC(Maintenance_Mode.OIT_Status) ][OTE(DO_Local_1.15) ,OTE(DO_L_1_15_Feed_Pump_Light_Out) ];
   16: [XIC(DO_R_3_0_Pure_Steam_Temp_Control_YV_4110.Activate) XIO(Maintenance_Mode.OIT_Status) ,XIC(DO_R_3_0_Pure_Steam_Temp_Control_YV_4110.Maint_Latch.OIT_Status) XIC(Maintenance_Mode.OIT_Status) ][OTE(DO_Remote_3.0) ,OTE(DO_R_3_0_Pure_Steam_Control_Valve_Out) ];
   17: [XIC(DO_R_3_1_Primary_Level_Control_YV_4760.Activate) XIO(Maintenance_Mode.OIT_Status) ,XIC(DO_R_3_1_Primary_Level_Control_YV_4760.Maint_Latch.OIT_Status) XIC(Maintenance_Mode.OIT_Status) ][OTE(DO_Remote_3.1) ,OTE(DO_R_3_1_Pri_Level_Valve_Out) ];
   18: [XIC(DO_R_3_2_Secondary_Level_Control_YV_4770.Activate) XIO(Maintenance_Mode.OIT_Status) ,XIC(DO_R_3_2_Secondary_Level_Control_YV_4770.Maint_Latch.OIT_Status) XIC(Maintenance_Mode.OIT_Status) ][OTE(DO_Remote_3.2) ,OTE(DO_R_3_2_Sec_Level_Valve_Out) ];
   19: [XIC(DO_R_3_3_Coolant_Shutoff_FCV_3025.Activate) XIO(Maintenance_Mode.OIT_Status) ,XIC(DO_R_3_3_Coolant_Shutoff_FCV_3025.Maint_Latch.OIT_Status) XIC(Maintenance_Mode.OIT_Status) ][OTE(DO_Remote_3.3) ,OTE(DO_R_3_3_Coolant_Valve_Out) ];
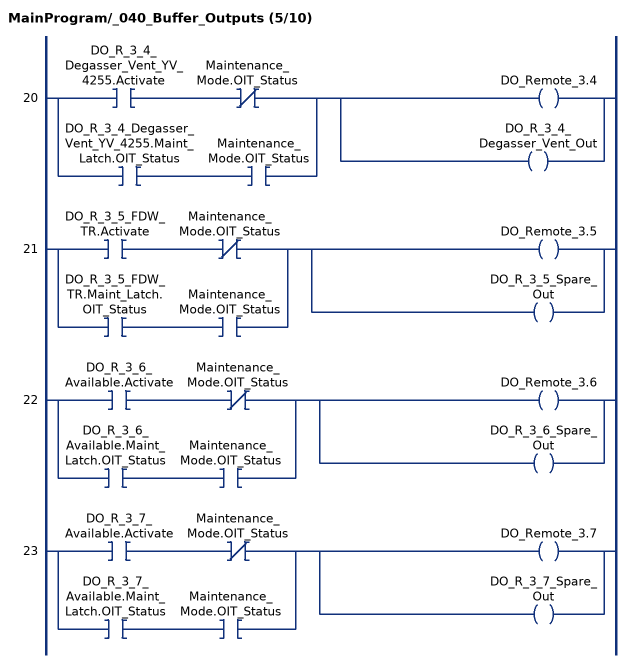
   20: [XIC(DO_R_3_4_Degasser_Vent_YV_4255.Activate) XIO(Maintenance_Mode.OIT_Status) ,XIC(DO_R_3_4_Degasser_Vent_YV_4255.Maint_Latch.OIT_Status) XIC(Maintenance_Mode.OIT_Status) ][OTE(DO_Remote_3.4) ,OTE(DO_R_3_4_Degasser_Vent_Out) ];
   21: [XIC(DO_R_3_5_FDW_TR.Activate) XIO(Maintenance_Mode.OIT_Status) ,XIC(DO_R_3_5_FDW_TR.Maint_Latch.OIT_Status) XIC(Maintenance_Mode.OIT_Status) ][OTE(DO_Remote_3.5) ,OTE(DO_R_3_5_Spare_Out) ];
   22: [XIC(DO_R_3_6_Available.Activate) XIO(Maintenance_Mode.OIT_Status) ,XIC(DO_R_3_6_Available.Maint_Latch.OIT_Status) XIC(Maintenance_Mode.OIT_Status) ][OTE(DO_Remote_3.6) ,OTE(DO_R_3_6_Spare_Out) ];
   23: [XIC(DO_R_3_7_Available.Activate) XIO(Maintenance_Mode.OIT_Status) ,XIC(DO_R_3_7_Available.Maint_Latch.OIT_Status) XIC(Maintenance_Mode.OIT_Status) ][OTE(DO_Remote_3.7) ,OTE(DO_R_3_7_Spare_Out) ];
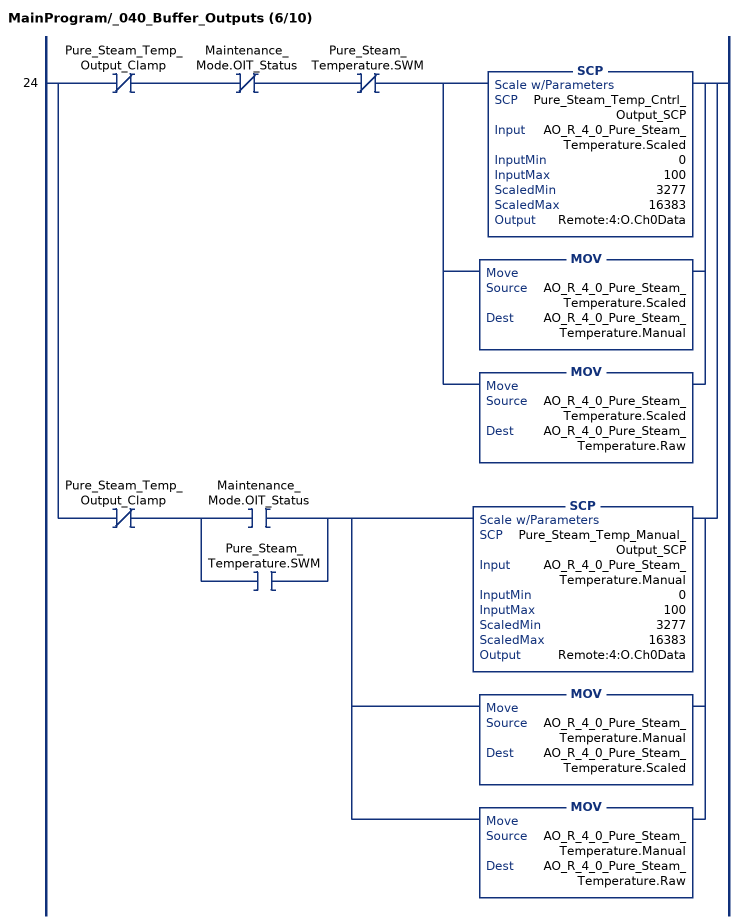
   24: [XIO(Pure_Steam_Temp_Output_Clamp) XIO(Maintenance_Mode.OIT_Status) XIO(Pure_Steam_Temperature.SWM) [SCP(Pure_Steam_Temp_Cntrl_Output_SCP,AO_R_4_0_Pure_Steam_Temperature.Scaled,0,100,3277,16383,Remote:4:O.Ch0Data) ,MOV(AO_R_4_0_Pure_Steam_Temperature.Scaled,AO_R_4_0_Pure_Steam_Temperature.Manual) ,MOV(AO_R_4_0_Pure_Steam_Temperature.Scaled,AO_R_4_0_Pure_Steam_Temperature.Raw) ] ,XIO(Pure_Steam_Temp_Output_Clamp) [XIC(Maintenance_Mode.OIT_Status) ,XIC(Pure_Steam_Temperature.SWM) ] [SCP(Pure_Steam_Temp_Manual_Output_SCP,AO_R_4_0_Pure_Steam_Temperature.Manual,0,100,3277,16383,Remote:4:O.Ch0Data) ,MOV(AO_R_4_0_Pure_Steam_Temperature.Manual,AO_R_4_0_Pure_Steam_Temperature.Scaled) ,MOV(AO_R_4_0_Pure_Steam_Temperature.Manual,AO_R_4_0_Pure_Steam_Temperature.Raw) ] ];
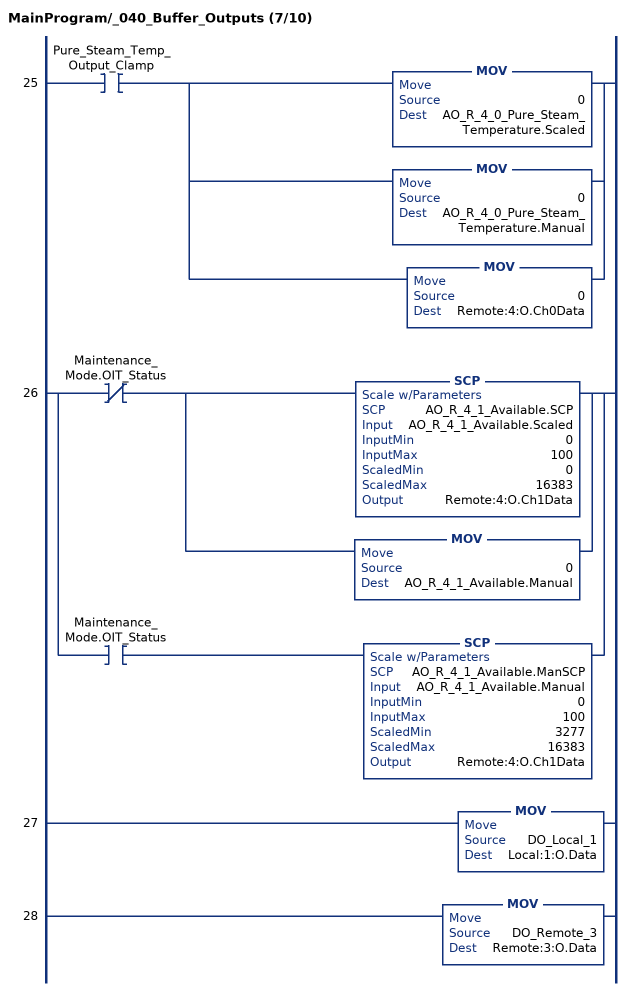
   25: XIC(Pure_Steam_Temp_Output_Clamp)[MOV(0,AO_R_4_0_Pure_Steam_Temperature.Scaled) ,MOV(0,AO_R_4_0_Pure_Steam_Temperature.Manual) ,MOV(0,Remote:4:O.Ch0Data) ];
   26: [XIO(Maintenance_Mode.OIT_Status) [SCP(AO_R_4_1_Available.SCP,AO_R_4_1_Available.Scaled,0,100,0,16383,Remote:4:O.Ch1Data) ,MOV(0,AO_R_4_1_Available.Manual) ] ,XIC(Maintenance_Mode.OIT_Status) SCP(AO_R_4_1_Available.ManSCP,AO_R_4_1_Available.Manual,0,100,3277,16383,Remote:4:O.Ch1Data) ];
   27: MOV(DO_Local_1,Local:1:O.Data);
   28: MOV(DO_Remote_3,Remote:3:O.Data);
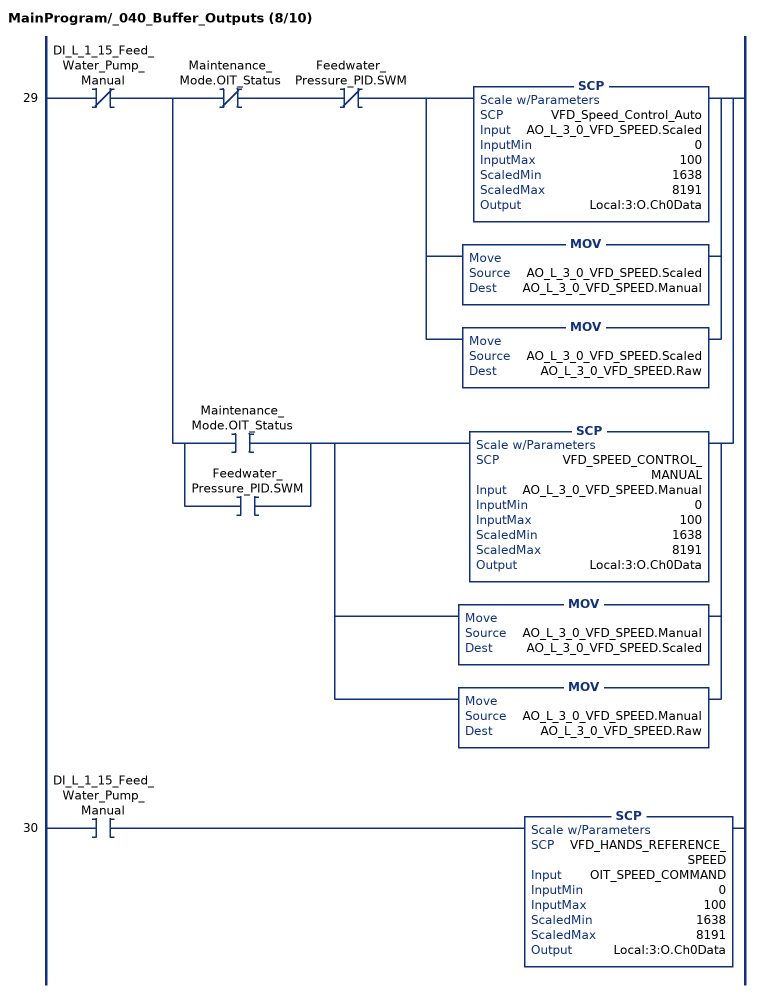
   29: XIO(DI_L_1_15_Feed_Water_Pump_Manual)[XIO(Maintenance_Mode.OIT_Status) XIO(Feedwater_Pressure_PID.SWM) [SCP(VFD_Speed_Control_Auto,AO_L_3_0_VFD_SPEED.Scaled,0,100,1638,8191,Local:3:O.Ch0Data) ,MOV(AO_L_3_0_VFD_SPEED.Scaled,AO_L_3_0_VFD_SPEED.Manual) ,MOV(AO_L_3_0_VFD_SPEED.Scaled,AO_L_3_0_VFD_SPEED.Raw) ] ,[XIC(Maintenance_Mode.OIT_Status) ,XIC(Feedwater_Pressure_PID.SWM) ] [SCP(VFD_SPEED_CONTROL_MANUAL,AO_L_3_0_VFD_SPEED.Manual,0,100,1638,8191,Local:3:O.Ch0Data) ,MOV(AO_L_3_0_VFD_SPEED.Manual,AO_L_3_0_VFD_SPEED.Scaled) ,MOV(AO_L_3_0_VFD_SPEED.Manual,AO_L_3_0_VFD_SPEED.Raw) ] ];
   30: XIC(DI_L_1_15_Feed_Water_Pump_Manual)SCP(VFD_HANDS_REFERENCE_SPEED,OIT_SPEED_COMMAND,0,100,1638,8191,Local:3:O.Ch0Data);
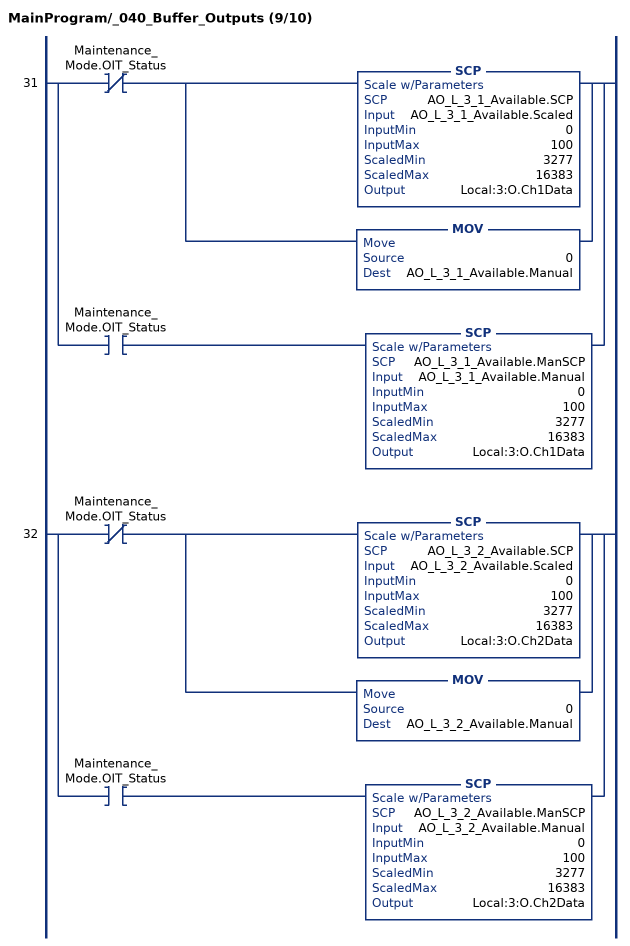
   31: [XIO(Maintenance_Mode.OIT_Status) [SCP(AO_L_3_1_Available.SCP,AO_L_3_1_Available.Scaled,0,100,3277,16383,Local:3:O.Ch1Data) ,MOV(0,AO_L_3_1_Available.Manual) ] ,XIC(Maintenance_Mode.OIT_Status) SCP(AO_L_3_1_Available.ManSCP,AO_L_3_1_Available.Manual,0,100,3277,16383,Local:3:O.Ch1Data) ];
   32: [XIO(Maintenance_Mode.OIT_Status) [SCP(AO_L_3_2_Available.SCP,AO_L_3_2_Available.Scaled,0,100,3277,16383,Local:3:O.Ch2Data) ,MOV(0,AO_L_3_2_Available.Manual) ] ,XIC(Maintenance_Mode.OIT_Status) SCP(AO_L_3_2_Available.ManSCP,AO_L_3_2_Available.Manual,0,100,3277,16383,Local:3:O.Ch2Data) ];
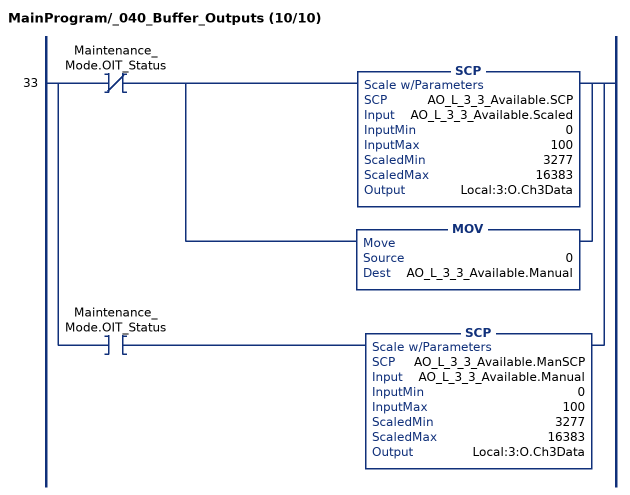
   33: [XIO(Maintenance_Mode.OIT_Status) [SCP(AO_L_3_3_Available.SCP,AO_L_3_3_Available.Scaled,0,100,3277,16383,Local:3:O.Ch3Data) ,MOV(0,AO_L_3_3_Available.Manual) ] ,XIC(Maintenance_Mode.OIT_Status) SCP(AO_L_3_3_Available.ManSCP,AO_L_3_3_Available.Manual,0,100,3277,16383,Local:3:O.Ch3Data) ];
END_ROUTINE
